(* IEC 61131-3 sources: stratumak/src/stmak/internal/modcompile/st/testdata/thirdparty/ironplc, 21 files *)

(* ---- first_steps_data_type_decl.st ---- *)
TYPE
  LOGLEVEL : (CRITICAL, WARNING, INFO, DEBUG) := INFO;
END_TYPE

(* ---- strings.st ---- *)
TYPE
   TEXT_EXTENDED : STRING [1] := '�';
END_TYPE

(* ---- array.st ---- *)
FUNCTION fun:BOOL

VAR_INPUT
    var1: INT;
    pt: ARRAY[1..8] OF INT;
END_VAR

var1 := var1 + pt[i];

END_FUNCTION

(* ---- array_in_function_var.st ---- *)
FUNCTION MY_FUNC : BOOL

VAR_INPUT
    x : INT;
END_VAR

VAR
    stack : ARRAY[1..32] OF UINT;
END_VAR

stack[1] := INT_TO_UINT(x);
MY_FUNC := TRUE;

END_FUNCTION

(* ---- array_of_string.st ---- *)
FUNCTION fun:BOOL

VAR_INPUT
    names: ARRAY[1..3] OF STRING[10];
END_VAR

fun := TRUE;

END_FUNCTION

(* ---- c_style_block_comment.st ---- *)
FUNCTION MY_FUNC : INT
VAR_INPUT
    x : INT;
END_VAR
    /* This is a C-style block comment */
    MY_FUNC := x;
END_FUNCTION

(* ---- empty_var_block.st ---- *)
FUNCTION myFunc : INT
VAR_INPUT
    x : INT;
END_VAR
VAR
END_VAR
    myFunc := x;
END_FUNCTION

(* ---- expressions.st ---- *)
FUNCTION fun:BOOL

VAR_INPUT
    var1: BYTE;
END_VAR

IF var1 < BYTE#32 THEN
	var1 := 1;
END_IF;

var1 := NOT (var3 OR var3);

var1 := FUNC_NAME(var1,'  ');

var1 := - 1 + 2 * 3 - 4 / 6 MOD 7 ** 8;

var1 := 1 >= 2 <= 3 <> 4 XOR 5;

IF var1 > t#1s THEN
    var1 := 1;
END_IF;

END_FUNCTION

(* ---- first_steps_func_avg_val.st ---- *)
FUNCTION AverageVal : REAL
    VAR_INPUT
    Cnt1 : INT;
    Cnt2 : INT;
    Cnt3 : INT;
    Cnt4 : INT;
    Cnt5 : INT;
  END_VAR
    VAR
    InputsNumber : REAL := 5.1;
  END_VAR
    AverageVal := INT_TO_REAL(Cnt1+Cnt2+Cnt3+Cnt4+Cnt5)/InputsNumber;
    END_FUNCTION

(* ---- inout_var_decl.st ---- *)
FUNCTION FUNC:UINT
    VAR_IN_OUT
        E : REAL;
        RNG : INT (1..2);
        ARR : ARRAY [0..3] OF INT;
    END_VAR

    array_avg := array_avg + arr[idx][idx];

END_FUNCTION

(* ---- input_var_decl.st ---- *)
FUNCTION FUNC:UINT
    VAR_INPUT
        E : REAL;
        PI, G : BOOL R_EDGE;
    END_VAR

    array_avg := array_avg + arr[idx][idx];

END_FUNCTION

(* ---- nested.st ---- *)
FUNCTION fun:BOOL

VAR_INPUT
    var1: BYTE;
END_VAR

array_avg := array_avg + arr[idx][idx];

END_FUNCTION

(* ---- comment.st ---- *)
(* COMMENT *)
FUNCTION_BLOCK BLOCK
    (* MULTI-LINE
       COMMENT *)
    VAR_INT := 10;
END_FUNCTION_BLOCK

(* ---- conditional.st ---- *)
FUNCTION_BLOCK BLOCK

    IF NOT VAR1 AND VAR1 THEN
        VAR1 := 1;
    ELSIF NOT VAR1 AND VAR1 THEN
        VAR1 := 1;
    END_IF;

END_FUNCTION_BLOCK

(* ---- first_steps_function_block_logger.st ---- *)
FUNCTION_BLOCK LOGGER
  VAR_INPUT
    TRIG : BOOL;
    MSG : STRING;
    LEVEL : LOGLEVEL := INFO;
  END_VAR
  VAR
    TRIG0 : BOOL;
  END_VAR

  IF TRIG AND NOT TRIG0 THEN

  END_IF;
  TRIG0:=TRIG;
END_FUNCTION_BLOCK

(* ---- if.st ---- *)
FUNCTION_BLOCK Error
    IF TRUE THEN
        Error := TRUE;
    END_IF
    IF TRUE THEN
        Error := TRUE;
    END_IF
END_FUNCTION_BLOCK

(* ---- literal.st ---- *)
FUNCTION_BLOCK BLOCK
    VAR
        REAL_WITH_TYPE: REAL := LREAL#11.0;
        BOOL_WITH_TYPE_TRUE: BOOL := BOOL#TRUE;
        TOD_WITH_VALUE_INTEGRAL: TIME_OF_DAY := TIME_OF_DAY#14:30:20;
        DATE_WITH_VALUE: DATE := DATE#2024-01-20;
        DATE_AND_TIME_WITH_VALUE: DATE_AND_TIME := DATE_AND_TIME#2024-01-20-15:30:22;
    END_VAR
    REAL_WITH_TYPE := 10;
END_FUNCTION_BLOCK

(* ---- textual.st ---- *)
FUNCTION_BLOCK BLOCK
    NUM_INT := 10;
    NUM_FLOAT := 10.0;

    IF NUM1 < NUM2 THEN
        NUM1 := 1;
    ELSIF NUM2 = NUM3 THEN
        NUM1 := 2;
    ELSE
        NUM1 := 3;
    END_IF;

    CASE EXPR_WITH_ELSE OF
    VAL1: (* empty *);
    VAL2: NUM1 := 1;
    ELSE NUM2 := 2;
    END_CASE;

    CASE EXPR_NO_ELSE OF
    VAL1: (* empty *);
    VAL2: NUM1 := 1;
    END_CASE;

    FOR VAL1 := 1 TO 10 BY 1 DO
       VAL2 := VAL1;
    END_FOR;

    WHILE VAL1 = 1 DO
        VAL2 := VAL1;
    END_WHILE;

    REPEAT
        VAL2 := VAL1;
    UNTIL VAL2 = 2
    END_REPEAT;

END_FUNCTION_BLOCK

(* ---- var_temp.st ---- *)
FUNCTION my_func : DINT
  VAR_INPUT
    a : DINT;
  END_VAR
  VAR_TEMP
    temp : DINT;
  END_VAR
  temp := a * 2;
  my_func := temp;
END_FUNCTION

FUNCTION_BLOCK my_fb
  VAR_TEMP
    t : INT;
  END_VAR
  t := 42;
END_FUNCTION_BLOCK

(* ---- first_steps_program.st ---- *)
PROGRAM plc_prg
  VAR_INPUT
    Reset : BOOL;
  END_VAR
  VAR_OUTPUT
    Cnt1 : INT;
    Cnt2 : INT;
    Cnt3 : INT;
    Cnt4 : INT;
    Cnt5 : INT;
  END_VAR
  VAR
    CounterST0 : CounterST;
    CounterFBD0 : CounterFBD;
    CounterSFC0 : CounterSFC;
    CounterIL0 : CounterIL;
    CounterLD0 : CounterLD;
    AVCnt : REAL;
    _TMP_AverageVal17_OUT : REAL;
  END_VAR

  CounterST0(Reset := Reset);
  Cnt1 := CounterST0.OUT;
  _TMP_AverageVal17_OUT := AverageVal(Cnt1, Cnt2, Cnt3, Cnt4, Cnt5);
  AVCnt := _TMP_AverageVal17_OUT;
  CounterFBD0(Reset := Reset);
  Cnt2 := CounterFBD0.OUT;
  CounterSFC0(Reset := Reset);
  Cnt3 := CounterSFC0.OUT;
  CounterIL0(Reset := Reset);
  Cnt4 := CounterIL0.OUT;
  CounterLD0(Reset := Reset);
  Cnt5 := CounterLD0.Out;
END_PROGRAM

(* ---- steel_thread.st ---- *)
PROGRAM main
  VAR
    x : INT;
    y : INT;
  END_VAR
  x := 10;
  y := x + 32;
END_PROGRAM
